(* IEC 61131-3 sources: codesys-framework/txt/application/WeVe Core (library)/10 Mode/ModeRequest/I_ModeRequest, 6 files *)

(* ---- ResetEvents.method.st ---- *)
METHOD ResetEvents : BOOL
VAR_INPUT
END_VAR

(* ---- ResetMachine.method.st ---- *)
METHOD ResetMachine : BOOL
VAR_INPUT
END_VAR

(* ---- ResetSafety.method.st ---- *)
METHOD ResetSafety : BOOL
VAR_INPUT
END_VAR

(* ---- StartRequest.method.st ---- *)
METHOD StartRequest : BOOL
VAR_INPUT
END_VAR

(* ---- StopRequest.method.st ---- *)
METHOD StopRequest : BOOL
VAR_INPUT
END_VAR

(* ---- UserRequest.method.st ---- *)
METHOD UserRequest : BOOL
VAR_INPUT
	nRequest	: UINT;
	pData		: POINTER TO ARRAY [0..255] OF BYTE := 0;
	pSize		: ULINT := 0;
END_VAR
